// TIA Portal V20 export
TYPE "WT2_Pf_Status_UDT"
   STRUCT
      iHandshake : Int;
      Datum : Array[0..9] of Char;
      Zeit : Array[0..7] of Char;
      SwVersion : Array[0..7] of Char;
      Fehler : Struct
         bE0000_KonfigFehler : Bool;
         bE0001_IOZuweisungUnvollst : Bool;
         bE0002_Reserviert : Bool;
         bE0003_Reserviert : Bool;
         bE0004_FehlerIOKomm : Bool;
         bE0005_FehlerKabelbruch : Bool;
         bE0006_FehlerIOHWKonfig : Bool;
         bE0007_Reserviert : Bool;
         bE0008_Reserviert : Bool;
         bE0009_Reserviert : Bool;
         bE0010_Reserviert : Bool;
         bE0011_Reserviert : Bool;
         bE0012_Reserviert : Bool;
         bE0013_Reserviert : Bool;
         bE0014_Reserviert : Bool;
         bE0015_Reserviert : Bool;
         bE0016_Reserviert : Bool;
         b301_Reserve : Bool;
         b302_Reserve : Bool;
         b303_Reserve : Bool;
         b304_Reserve : Bool;
         b305_Reserve : Bool;
         b306_Reserve : Bool;
         b307_Reserve : Bool;
         by31_Reserve : Byte;
      END_STRUCT;
      Alarm : Struct
         bA1000_Reserviert : Bool;
         bA1001_Reserviert : Bool;
         bA1002_Reserviert : Bool;
         bA1003_Reserviert : Bool;
         bA1004_Reserviert : Bool;
         bA1005_AlarmKabelbruch : Bool;
         bA1006_Reserviert : Bool;
         bA1007_AlarmFeldbus : Bool;
         bA1008_ZugriffsfehlerCFKarte : Bool;
         bA1009_MZeitMasterAktiv : Bool;
         bA1010_FehlerInitSteuerkomm : Bool;
         bA1011_AlarmFBStandbyMasterAktiv : Bool;
         bA1012_Reserviert : Bool;
         bA1013_AlarmFehlerIOModul : Bool;
         bA1014_AlarmFehlerIOModulAnz : Bool;
         bA1015_AlarmCPUTempZuHoch : Bool;
         bA1016_AlarmCPUAuslZuHoch : Bool;
         b341_Reserve : Bool;
         b342_Reserve : Bool;
         b343_Reserve : Bool;
         b344_Reserve : Bool;
         b345_Reserve : Bool;
         b346_Reserve : Bool;
         b347_Reserve : Bool;
         by35_Reserve : Byte;
      END_STRUCT;
      Zustand : Struct
         bFehlerzustandAktiv : Bool;
         bAlarmzustandAktiv : Bool;
         bSystemMeldungAktiv : Bool;
         bSeviceMeldungAktiv : Bool;
         bStopManuell : Bool;
         bStopAuto : Bool;
         bStopExtern : Bool;
         bBetriebAuto : Bool;
         bBetriebManuell : Bool;
         bAnlaufAuto : Bool;
         bAnlaufManuell : Bool;
         bManuellStoppen : Bool;
         b374_Reserve : Bool;
         b375_Reserve : Bool;
         b376_Reserve : Bool;
         b377_Reserve : Bool;
         by38_Reserve : Byte;
         bSystemMeldungKonfigUmschaltung : Bool;
         b391_Reserve : Bool;
         b392_Reserve : Bool;
         b393_Reserve : Bool;
         b394_Reserve : Bool;
         b395_Reserve : Bool;
         b396_Reserve : Bool;
         b397_Reserve : Bool;
         by40_Reserve : Byte;
         by41_Reserve : Byte;
         by42_Reserve : Byte;
         by43_Reserve : Byte;
      END_STRUCT;
      DigIn : Struct
         bKonfigSatzBit0 : Bool;
         bKonfigSatzBit1 : Bool;
         bFreigabeTempRegler : Bool;
         bFreigabeZweipunktRegler1 : Bool;
         bFreigabeZweipunktRegler2 : Bool;
         bFreigabeZweipunktregler3 : Bool;
         bFreigabeZweipunktregler4 : Bool;
         bFreigabePIRegler1 : Bool;
         bFreigabePIRegler2 : Bool;
         bFreigabePIRegler3 : Bool;
         bFreigabePIRegler4 : Bool;
         b453_Reserve : Bool;
         b454_Reserve : Bool;
         b455_Reserve : Bool;
         b456_Reserve : Bool;
         b457_Reserve : Bool;
         by46_Reserve : Byte;
         by47_Reserve : Byte;
      END_STRUCT;
      DigOut : Struct
         bFehler : Bool;
         bAlarm : Bool;
         bTemperaturregler : Bool;
         bZweipunktrelger1 : Bool;
         bZweipunktrelger2 : Bool;
         bZweipunktregler3 : Bool;
         bZweipunktregler4 : Bool;
         b487_Reserve : Bool;
         by49_Reserve : Byte;
         by50_Reserve : Byte;
         by51_Reserve : Byte;
      END_STRUCT;
      iKonfigSatz : Int;
      rReserveReal : Array[0..9] of Real;
      byReserveByte : Array[0..1] of Byte;
   END_STRUCT;
END_TYPE
